(* IEC 61131-3 sources: ZPLC/packages/zplc-ide/projects/edge_counter/src, 1 file *)

(* ---- EdgeCounter.st ---- *)
(*
 * Edge Counter - count three pulses, then hold CountReached until Reset.
 *
 * CTU counts rising edges of CU on its own: it keeps CU from the previous scan and adds one only on a FALSE-to-TRUE
 * change. A pulse therefore counts once however many scans it stays high, and PulseInput can be wired straight to CU.
 * An R_TRIG in front of CTU would only turn the same edge into a one-scan pulse that CTU then edge-detects a second time.
 *
 * Reset sets the count to 0 and CountReached to FALSE. CTU keeps watching CU while Reset is TRUE, as the IEC definition
 * does, so a pulse that rises during Reset is not counted when Reset is released, even if it is still high. Only a new
 * rising edge after that counts: a pulse that arrives while Reset is held is lost.
 *)

PROGRAM EdgeCounter

VAR_INPUT
    PulseInput AT %I0.0 : BOOL;
    Reset AT %I0.1 : BOOL;
END_VAR

VAR
    Count : CTU;                    (* up counter: Count.CV is the count so far *)
END_VAR

VAR_OUTPUT
    CountReached AT %Q0.0 : BOOL;   (* TRUE once Count.CV has reached the preset *)
END_VAR

Count(CU := PulseInput, R := Reset, PV := 3);
CountReached := Count.Q;

END_PROGRAM
